Fanuc KAREL source: KT00517.KL

PROGRAM KT00517
%NOLOCKGROUP
VAR
  P1: XYZWPREXT
  P2: POSITION
  OUT: JOINTPOS
BEGIN
  P1.X = 1.0
  OUT = P1 : P2
END KT00517
